(* IEC 61131-3 sources: canworks/examples/openplc-fuxa/pous/programs, 3 files *)

(* ---- canworks_in.st ---- *)
PROGRAM canworks_in
  VAR
    i0  : WORD AT %IW100; (* cw_map_hash *)
    i1  : WORD AT %IW101; (* cw_map_hash_w1 *)
    i2  : WORD AT %IW102; (* cw_status *)
    i3  : WORD AT %IW103; (* cw_status_w1 *)
    i4  : WORD AT %IW104; (* cw_status_w2 *)
    i5  : WORD AT %IW105; (* cw_status_w3 *)
    i6  : WORD AT %IW106; (* rtd_temp1 *)
    i7  : WORD AT %IW107; (* rtd_temp2 *)
    i8  : WORD AT %IW108; (* rtd_AI2_Input_PV *)
    i9  : WORD AT %IW109; (* rtd_AI3_Input_PV *)
    i10 : WORD AT %IW110; (* dio_in0 *)
    i11 : WORD AT %IW111; (* dio_Read_analogue_input_1 *)
    i12 : WORD AT %IW112; (* dio_Read_analogue_input_2 *)
    i13 : WORD AT %IW113; (* can_bus_state *)
    i14 : WORD AT %IW114; (* rtd_ok *)
    i15 : WORD AT %IW115; (* rtd_emcy *)
    i16 : WORD AT %IW116; (* dio_state *)
    i17 : WORD AT %IW117; (* dio_emcy *)
    i18 : WORD AT %IW118; (* cw_live_list_field *)
    i19 : WORD AT %IW119; (* cw_live_list_field_w1 *)
    i20 : WORD AT %IW120; (* cw_live_list_field_w2 *)
    i21 : WORD AT %IW121; (* cw_live_list_field_w3 *)
    i22 : WORD AT %IW122; (* cw_live_list_field_w4 *)
    i23 : WORD AT %IW123; (* cw_live_list_field_w5 *)
    i24 : WORD AT %IW124; (* cw_live_list_field_w6 *)
    i25 : WORD AT %IW125; (* cw_live_list_field_w7 *)
    i26 : WORD AT %IW126; (* cw_sdo_bridge_response *)
    i27 : WORD AT %IW127; (* cw_sdo_bridge_response_w1 *)
    i28 : WORD AT %IW128; (* cw_sdo_bridge_response_w2 *)
    i29 : WORD AT %IW129; (* cw_sdo_bridge_response_w3 *)
    i30 : WORD AT %IW130; (* cw_sdo_bridge_response_w4 *)
    i31 : WORD AT %IW131; (* cw_sdo_bridge_response_w5 *)
    i32 : WORD AT %IW132; (* cw_sdo_bridge_response_w6 *)
  END_VAR
  VAR
    last_counter : WORD;
    moved        : BOOL;
    stale        : TON;
  END_VAR

(* Generated by canworks from canworks/canworks.json: do not edit, Save rewrites it. *)
moved := i3 <> last_counter;
last_counter := i3;
stale(IN := NOT moved, PT := T#300ms);
canworks.ok := i0 = WORD#16#54FD AND i1 = WORD#16#9749 AND NOT stale.Q;
canworks.bus_ok := canworks.ok AND (i5 AND WORD#16#0002) = WORD#0;
canworks.link[21] := WORD#16#0106 OR SEL(canworks.ok, WORD#0, WORD#1);
canworks.link[0] := i2;
canworks.link[1] := i3;
canworks.link[2] := i4;
canworks.link[3] := i5;
canworks.link[14] := i26;
canworks.link[15] := i27;
canworks.link[16] := i28;
canworks.link[17] := i29;
canworks.link[18] := i30;
canworks.link[19] := i31;
canworks.link[20] := i32;
canworks.link[25] := i18;
canworks.link[26] := i19;
canworks.link[27] := i20;
canworks.link[28] := i21;
canworks.link[29] := i22;
canworks.link[30] := i23;
canworks.link[31] := i24;
canworks.link[32] := i25;
canworks.can_bus_state := SEL(canworks.ok, USINT#0, WORD_TO_USINT((i13 AND WORD#16#00FF)));
canworks.can_master_state := SEL(canworks.ok, USINT#0, WORD_TO_USINT(SHR(i13, 8)));
canworks.rtd_ok := SEL(canworks.ok, FALSE, (i14 AND WORD#16#0100) <> WORD#0);
canworks.rtd_state := SEL(canworks.ok, USINT#0, WORD_TO_USINT((i14 AND WORD#16#00FF)));
canworks.rtd_emcy := SEL(canworks.ok, WORD#0, i15);
canworks.rtd_tpdo1_timeout := SEL(canworks.ok, FALSE, (i14 AND WORD#16#0200) <> WORD#0);
canworks.rtd_temp1 := WORD_TO_INT(i6);
canworks.rtd_temp2 := WORD_TO_INT(i7);
canworks.rtd_AI2_Input_PV := WORD_TO_INT(i8);
canworks.rtd_AI3_Input_PV := WORD_TO_INT(i9);
canworks.dio_ok := SEL(canworks.ok, FALSE, (i14 AND WORD#16#0400) <> WORD#0);
canworks.dio_state := SEL(canworks.ok, USINT#0, WORD_TO_USINT(SHR(i16, 8)));
canworks.dio_emcy := SEL(canworks.ok, WORD#0, i17);
canworks.dio_in0 := WORD_TO_USINT(SHR(i10, 8));
canworks.dio_in1 := WORD_TO_USINT((i10 AND WORD#16#00FF));
canworks.dio_Read_analogue_input_1 := WORD_TO_INT(i11);
canworks.dio_Read_analogue_input_2 := WORD_TO_INT(i12);

END_PROGRAM

(* ---- canworks_out.st ---- *)
PROGRAM canworks_out
  VAR
    q0  : WORD AT %QW100; (* cw_plc_link *)
    q1  : WORD AT %QW101; (* cw_plc_link_w1 *)
    q2  : WORD AT %QW102; (* cw_plc_link_w2 *)
    q3  : WORD AT %QW103; (* dio_out0 *)
    q4  : WORD AT %QW104; (* dio_Write_analogue_output_1 *)
    q5  : WORD AT %QW105; (* dio_Write_analogue_output_2 *)
    q6  : WORD AT %QW106; (* cw_control *)
    q7  : WORD AT %QW107; (* cw_control_w1 *)
    q8  : WORD AT %QW108; (* cw_control_w2 *)
    q9  : WORD AT %QW109; (* cw_sdo_bridge_request *)
    q10 : WORD AT %QW110; (* cw_sdo_bridge_request_w1 *)
    q11 : WORD AT %QW111; (* cw_sdo_bridge_request_w2 *)
    q12 : WORD AT %QW112; (* cw_sdo_bridge_request_w3 *)
    q13 : WORD AT %QW113; (* cw_sdo_bridge_request_w4 *)
    q14 : WORD AT %QW114; (* cw_sdo_bridge_request_w5 *)
    q15 : WORD AT %QW115; (* cw_sdo_bridge_request_w6 *)
  END_VAR

(* Generated by canworks from canworks/canworks.json: do not edit, Save rewrites it. *)
q3 := SHL((USINT_TO_WORD(canworks.dio_out0) AND WORD#16#00FF), 8) OR (USINT_TO_WORD(canworks.dio_out1) AND WORD#16#00FF);
q4 := INT_TO_WORD(canworks.dio_Write_analogue_output_1);
q5 := INT_TO_WORD(canworks.dio_Write_analogue_output_2);
q6 := canworks.link[4];
q7 := canworks.link[5];
q8 := canworks.link[6];
q9 := canworks.link[7];
q10 := canworks.link[8];
q11 := canworks.link[9];
q12 := canworks.link[10];
q13 := canworks.link[11];
q14 := canworks.link[12];
q15 := canworks.link[13];
(* PLC link header, last: running, then the map hash 0x54fd9749 *)
q1 := WORD#16#54FD;
q2 := WORD#16#9749;
q0 := WORD#1;

END_PROGRAM

(* ---- main.st ---- *)
(* The HMI's variables: FUXA reads and writes them by name over the
   project's OPC UA server (devices/servers/opcua.json). The CAN values
   come from the canworks variable list, which canworks_in fills before
   and canworks_out sends after this program in every scan. *)
PROGRAM main
  VAR
    temp1 : REAL;              (* temperature 1, degrees C *)
    temp2 : REAL;              (* temperature 2, degrees C *)
    limit : REAL := 25.0;      (* written by the HMI *)
    ack : BOOL;                (* written by the HMI; cleared after use *)
    run : BOOL := TRUE;        (* running light on, written by the HMI *)
    alarm : BOOL;
    light_ok : BOOL;
    canworks_ok : BOOL;        (* the bridge answers with this program's map *)
    bus_ok : BOOL;             (* and the CAN bus is up *)
    rtd_ok : BOOL;             (* node 5 operational *)
    dio_ok : BOOL;             (* node 6 operational *)
    dio_in0 : USINT;
    dio_in1 : USINT;
    dio_out0 : USINT;
    dio_out1 : USINT;
    manual_out0 : USINT;       (* bits 1-7 of dio_out0, written by the HMI *)
    manual_out1 : USINT;       (* dio_out1 while run is off, written by the HMI *)
    logic : PLANT_LOGIC;
  END_VAR

  canworks_ok := canworks.ok;
  bus_ok := canworks.bus_ok;
  rtd_ok := canworks.rtd_ok;
  dio_ok := canworks.dio_ok;
  temp1 := INT_TO_REAL(canworks.rtd_temp1) / 10.0;
  temp2 := INT_TO_REAL(canworks.rtd_temp2) / 10.0;
  dio_in0 := canworks.dio_in0;
  dio_in1 := canworks.dio_in1;

  logic(VALID := canworks_ok AND rtd_ok, TEMP := temp1, LIMIT := limit, ACK := ack, RUN := run,
        DIO_IN1 := dio_in1, MANUAL_OUT0 := manual_out0, MANUAL_OUT1 := manual_out1);
  alarm := logic.ALARM;
  light_ok := logic.LIGHT_OK;
  dio_out0 := logic.DIO_OUT0;
  dio_out1 := logic.DIO_OUT1;
  ack := FALSE;

  canworks.dio_out0 := dio_out0;
  canworks.dio_out1 := dio_out1;
END_PROGRAM
